// TIA Portal V20 export
FUNCTION_BLOCK "PR_IRVisionCheckSeq_Soft2.0 1_workflow_93eeda"   // FB47, LAD
{ S7_Optimized_Access := 'TRUE' }
// stored: MemoryReserve 100, SetENOAutomatically false
   VAR_INPUT
      iAutoRunning : Bool;
      iFaultReset : Bool;
      iIRMesaureProbeDown : Bool;
      iIRMesaureProbeUp : Bool;
      iIndexCylHome : Bool;
      iIndexProbeOut : Bool;
      iInspectionOver : Bool;
      iManualEntryConfirm : Bool;
      iMesauringOver : Bool;
      iProbeCylHome : Bool;
      iRFIDReadError : Bool;
      iRFIDReadOver : Bool;
      iReject : Bool;
      iReset_fault : Bool;
      iRetry : Bool;
      iRetryCount : Int;
      iSstMode : Bool;
      iSstPB : Bool;
      iStartFrmFibroseq : Bool;
   END_VAR
   VAR_OUTPUT
      qCameraLight : Bool;
      qError : Array[0..9] of Bool;
      qIRProbeDown : Bool;
      qIRProbeUp : Bool;
      qIRVisionCheckOver : Bool;
      qIndexProbeIn : Bool;
      qIndexProbeOut : Bool;
      qMessage : Array[0..9] of Bool;
   END_VAR
   VAR
      c20_ChkRecoveryStatus_T1 : Bool;
      c20_ChkRecoveryStatus_T2 : Bool;
      c20_ChkRecoveryStatus_T3 : Bool;
      c20_ChkRecoveryStatus_T4 : Bool;
      c22_WtRFIDReadOver_T1 : Bool;
      c22_WtRFIDReadOver_T2 : Bool;
      c23_ChkRetryCountOver_T1 : Bool;
      c23_ChkRetryCountOver_T2 : Bool;
      c24_WtOperatorDecisionRead_T1 : Bool;
      c24_WtOperatorDecisionRead_T2 : Bool;
      c25_ChkPartWorkable_T1 : Bool;
      c25_ChkPartWorkable_T2 : Bool;
      c91_WtRFIDWriteOver_T1 : Bool;
      c91_WtRFIDWriteOver_T2 : Bool;
      c92_ChkWriteRetryCountOver_T1 : Bool;
      c92_ChkWriteRetryCountOver_T2 : Bool;
      c93_WtOperatorDecisionWrite_T1 : Bool;
      c93_WtOperatorDecisionWrite_T2 : Bool;
      StateNo : Int;
      s100_WtStartLow : Bool;
      s100_WtStartLow_T1 : Bool;
      s10_WtStartFrmFibroSeq : Bool;
      s10_WtStartFrmFibroSeq_T1 : Bool;
      s1_WtResetRel : Bool;
      s1_WtResetRel_T1 : Bool;
      s20_ChkRecoveryStatus : Bool;
      s20_ChkRecoveryStatus_T1 : Bool;
      s20_ChkRecoveryStatus_T2 : Bool;
      s20_ChkRecoveryStatus_T3 : Bool;
      s20_ChkRecoveryStatus_T4 : Bool;
      s21_WtProbeIndexCylHome : Bool;
      s21_WtProbeIndexCylHome_T1 : Bool;
      s22_WtRFIDReadOver : Bool;
      s22_WtRFIDReadOver_T1 : Bool;
      s22_WtRFIDReadOver_T2 : Bool;
      s23_ChkRetryCountOver : Bool;
      s23_ChkRetryCountOver_T1 : Bool;
      s23_ChkRetryCountOver_T2 : Bool;
      s24_WtOperatorDecisionRead : Bool;
      s24_WtOperatorDecisionRead_T1 : Bool;
      s24_WtOperatorDecisionRead_T2 : Bool;
      s25_ChkPartWorkable : Bool;
      s25_ChkPartWorkable_T1 : Bool;
      s25_ChkPartWorkable_T2 : Bool;
      s30_WtOperatorAck : Bool;
      s30_WtOperatorAck_T1 : Bool;
      s50_WtIRMeasureProbeAtTest : Bool;
      s50_WtIRMeasureProbeAtTest_T1 : Bool;
      s60_WtMeasurementOver : Bool;
      s60_WtMeasurementOver_T1 : Bool;
      s70_WtIRMeasureProbeUp : Bool;
      s70_WtIRMeasureProbeUp_T1 : Bool;
      s80_WtIndexingProbeOut : Bool;
      s80_WtIndexingProbeOut_T1 : Bool;
      s90_WtVisionInspectionOver : Bool;
      s90_WtVisionInspectionOver_T1 : Bool;
      s91_WtRFIDWriteOver : Bool;
      s91_WtRFIDWriteOver_T1 : Bool;
      s91_WtRFIDWriteOver_T2 : Bool;
      s92_ChkWriteRetryCountOver : Bool;
      s92_ChkWriteRetryCountOver_T1 : Bool;
      s92_ChkWriteRetryCountOver_T2 : Bool;
      s93_WtOperatorDecisionWrite : Bool;
      s93_WtOperatorDecisionWrite_T1 : Bool;
      s93_WtOperatorDecisionWrite_T2 : Bool;
      s94_WtAllSystemAtHome : Bool;
      s94_WtAllSystemAtHome_T1 : Bool;
      sAbnormalStatus : Bool;
      sIRInProgress : Bool;
      sPartWorkable : Bool;
      sRFReadRetryCount : Int;
      sRFWriteError : Bool;
      sRFWriteOver : Bool;
      sRFWriteRetryCount : Int;
      sSst : Bool;
      sSstPulse : Bool;
      sSstRise : Bool;
      sStWtResetRel : Bool;
      sStWtResetRel_T1 : Bool;
      sTimeouTime : TON_TIME;
      sVisionInProgress : Bool;
   END_VAR
   VAR_TEMP
      tOne : Bool;
   END_VAR
   VAR_TEMP   // added for the SCL form of the ladder/FBD networks
      _w1 : Bool;
   END_VAR
BEGIN

REGION Network 1
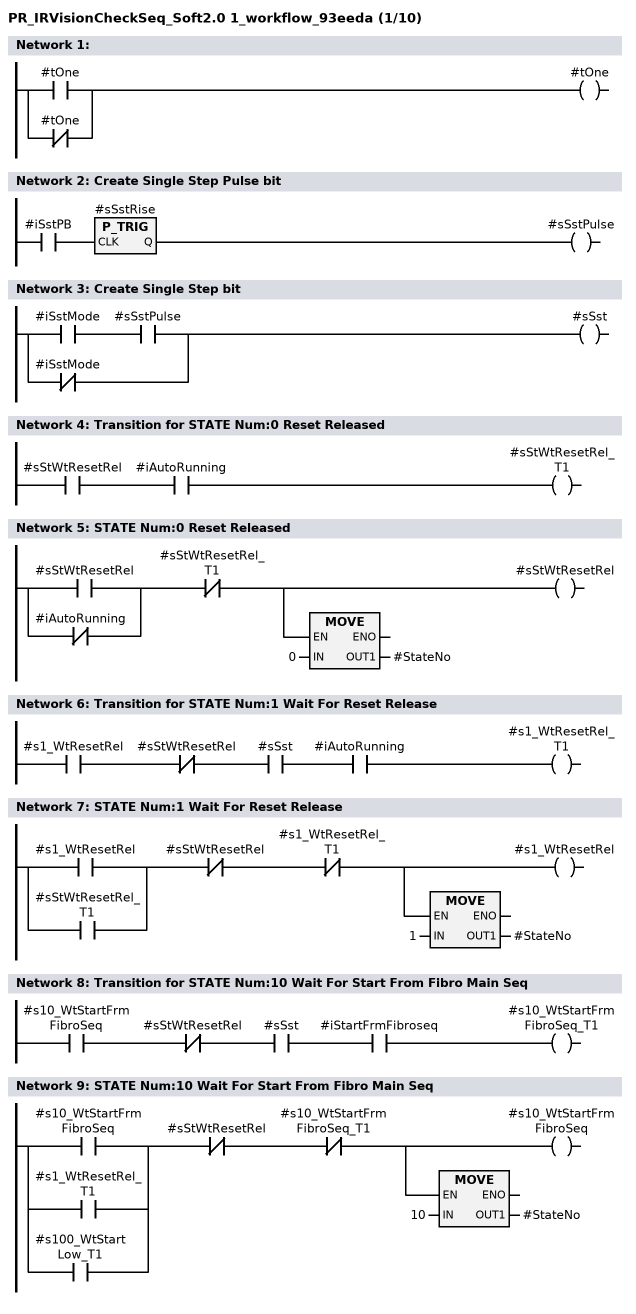
   RUNG wire#powerrail
      Contact( #tOne )
      wire#w1
      Coil( #tOne )
   END_RUNG
   RUNG wire#powerrail
      I_Contact( #tOne )
   END_RUNG wire#w1
   // the same network as SCL:
   #tOne := #tOne OR NOT #tOne;
END_REGION

REGION Network 2: Create Single Step Pulse bit
   RUNG wire#powerrail
      Contact( #iSstPB )
      P_Trig( #sSstRise )
      Coil( #sSstPulse )
   END_RUNG
   // the same network as SCL:
   #_w1 := #iSstPB AND NOT #sSstRise;   // rising edge
   #sSstRise := #iSstPB;
   #sSstPulse := #_w1;
END_REGION

REGION Network 3: Create Single Step bit
   RUNG wire#powerrail
      Contact( #iSstMode )
      Contact( #sSstPulse )
      wire#w1
      Coil( #sSst )
   END_RUNG
   RUNG wire#powerrail
      I_Contact( #iSstMode )
   END_RUNG wire#w1
   // the same network as SCL:
   #sSst := (#iSstMode AND #sSstPulse) OR NOT #iSstMode;
END_REGION

REGION Network 4: Transition for STATE Num:0 Reset Released
   RUNG wire#powerrail
      Contact( #sStWtResetRel )
      Contact( #iAutoRunning )
      Coil( #sStWtResetRel_T1 )
   END_RUNG
   // the same network as SCL:
   #sStWtResetRel_T1 := #sStWtResetRel AND #iAutoRunning;
END_REGION

REGION Network 5: STATE Num:0 Reset Released
   RUNG wire#powerrail
      Contact( #sStWtResetRel )
      wire#w1
      I_Contact( #sStWtResetRel_T1 )
      wire#w2
      Coil( #sStWtResetRel )
   END_RUNG
   RUNG wire#powerrail
      I_Contact( #iAutoRunning )
   END_RUNG wire#w1
   RUNG wire#w2
      { S7_GenerateENO := "TRUE" } Move(in := 0, out1 => #StateNo)
   END_RUNG
   // the same network as SCL:
   #sStWtResetRel := (#sStWtResetRel OR NOT #iAutoRunning) AND NOT #sStWtResetRel_T1;
   IF #sStWtResetRel THEN #StateNo := 0; END_IF;
END_REGION

REGION Network 6: Transition for STATE Num:1 Wait For Reset Release
   RUNG wire#powerrail
      Contact( #s1_WtResetRel )
      I_Contact( #sStWtResetRel )
      Contact( #sSst )
      Contact( #iAutoRunning )
      Coil( #s1_WtResetRel_T1 )
   END_RUNG
   // the same network as SCL:
   #s1_WtResetRel_T1 := #s1_WtResetRel AND NOT #sStWtResetRel AND #sSst AND #iAutoRunning;
END_REGION

REGION Network 7: STATE Num:1 Wait For Reset Release
   RUNG wire#powerrail
      Contact( #s1_WtResetRel )
      wire#w1
      I_Contact( #sStWtResetRel )
      I_Contact( #s1_WtResetRel_T1 )
      wire#w2
      Coil( #s1_WtResetRel )
   END_RUNG
   RUNG wire#powerrail
      Contact( #sStWtResetRel_T1 )
   END_RUNG wire#w1
   RUNG wire#w2
      { S7_GenerateENO := "TRUE" } Move(in := 1, out1 => #StateNo)
   END_RUNG
   // the same network as SCL:
   #s1_WtResetRel := (#s1_WtResetRel OR #sStWtResetRel_T1) AND NOT #sStWtResetRel AND NOT #s1_WtResetRel_T1;
   IF #s1_WtResetRel THEN #StateNo := 1; END_IF;
END_REGION

REGION Network 8: Transition for STATE Num:10 Wait For Start From Fibro Main Seq
   RUNG wire#powerrail
      Contact( #s10_WtStartFrmFibroSeq )
      I_Contact( #sStWtResetRel )
      Contact( #sSst )
      Contact( #iStartFrmFibroseq )
      Coil( #s10_WtStartFrmFibroSeq_T1 )
   END_RUNG
   // the same network as SCL:
   #s10_WtStartFrmFibroSeq_T1 := #s10_WtStartFrmFibroSeq AND NOT #sStWtResetRel AND #sSst AND #iStartFrmFibroseq;
END_REGION

REGION Network 9: STATE Num:10 Wait For Start From Fibro Main Seq
   RUNG wire#powerrail
      Contact( #s10_WtStartFrmFibroSeq )
      wire#w1
      I_Contact( #sStWtResetRel )
      I_Contact( #s10_WtStartFrmFibroSeq_T1 )
      wire#w2
      Coil( #s10_WtStartFrmFibroSeq )
   END_RUNG
   RUNG wire#powerrail
      Contact( #s1_WtResetRel_T1 )
   END_RUNG wire#w1
   RUNG wire#powerrail
      Contact( #s100_WtStartLow_T1 )
   END_RUNG wire#w1
   RUNG wire#w2
      { S7_GenerateENO := "TRUE" } Move(in := 10, out1 => #StateNo)
   END_RUNG
   // the same network as SCL:
   #s10_WtStartFrmFibroSeq := (#s10_WtStartFrmFibroSeq OR #s1_WtResetRel_T1 OR #s100_WtStartLow_T1) AND NOT #sStWtResetRel AND NOT #s10_WtStartFrmFibroSeq_T1;
   IF #s10_WtStartFrmFibroSeq THEN #StateNo := 10; END_IF;
END_REGION

REGION Network 10: Actions for STATE Num:10 Wait For Start From Fibro Main Seq
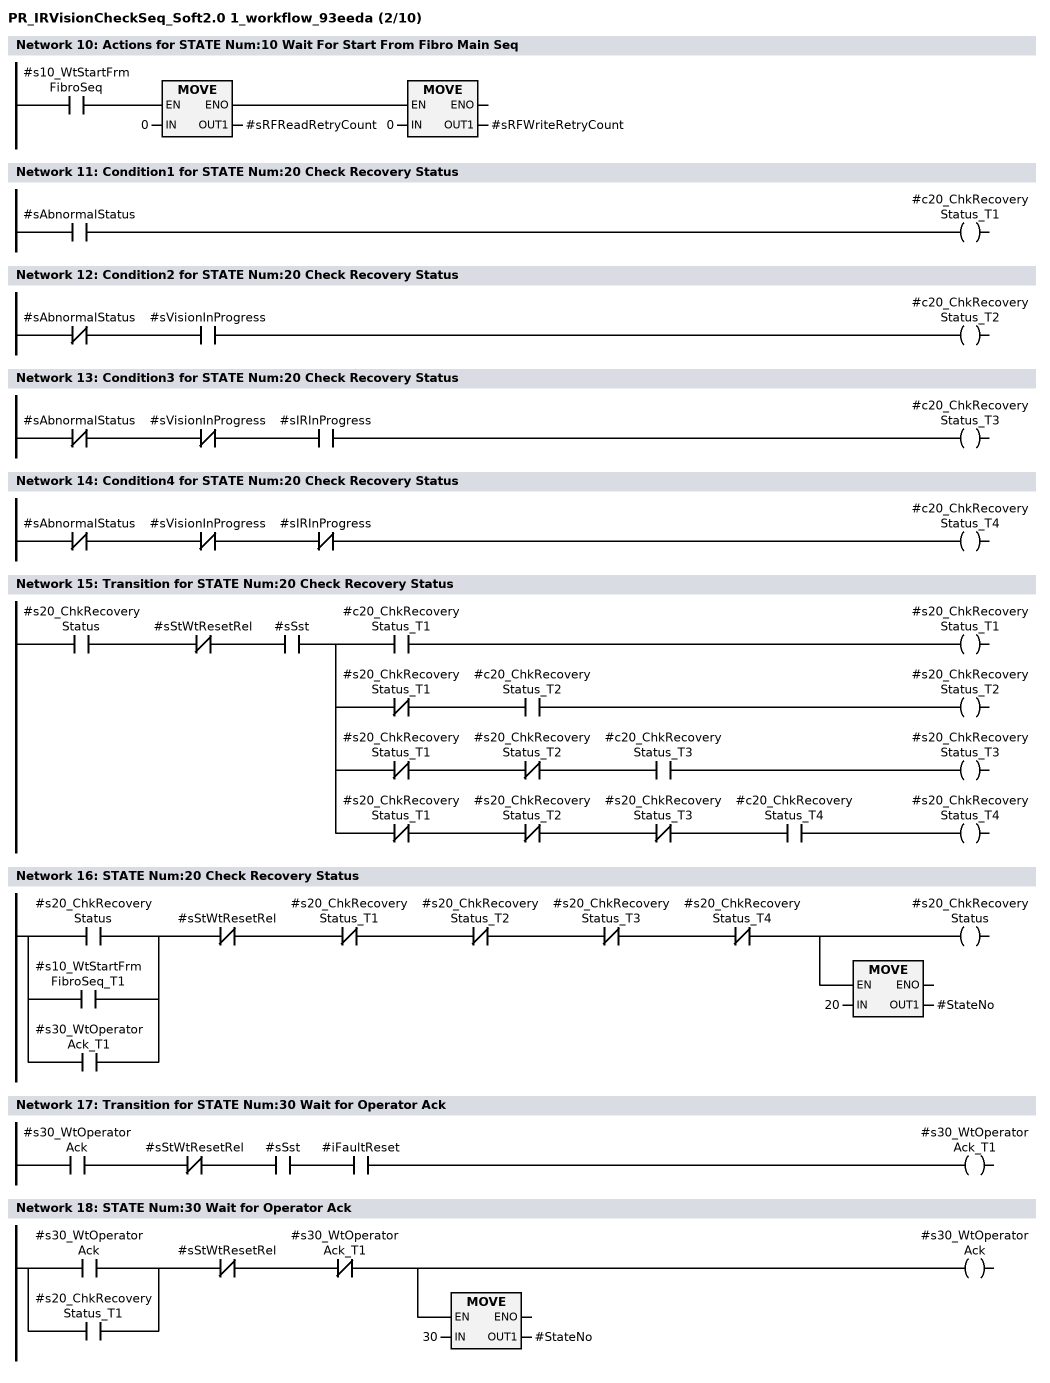
   RUNG wire#powerrail
      Contact( #s10_WtStartFrmFibroSeq )
      Move(in := 0, out1 => #sRFReadRetryCount)
      Move(in := 0, out1 => #sRFWriteRetryCount)
   END_RUNG
   // the same network as SCL:
   IF #s10_WtStartFrmFibroSeq THEN
       #sRFReadRetryCount := 0;
       #sRFWriteRetryCount := 0;
   END_IF;
END_REGION

REGION Network 11: Condition1 for STATE Num:20 Check Recovery Status
   RUNG wire#powerrail
      Contact( #sAbnormalStatus )
      Coil( #c20_ChkRecoveryStatus_T1 )
   END_RUNG
   // the same network as SCL:
   #c20_ChkRecoveryStatus_T1 := #sAbnormalStatus;
END_REGION

REGION Network 12: Condition2 for STATE Num:20 Check Recovery Status
   RUNG wire#powerrail
      I_Contact( #sAbnormalStatus )
      Contact( #sVisionInProgress )
      Coil( #c20_ChkRecoveryStatus_T2 )
   END_RUNG
   // the same network as SCL:
   #c20_ChkRecoveryStatus_T2 := NOT #sAbnormalStatus AND #sVisionInProgress;
END_REGION

REGION Network 13: Condition3 for STATE Num:20 Check Recovery Status
   RUNG wire#powerrail
      I_Contact( #sAbnormalStatus )
      I_Contact( #sVisionInProgress )
      Contact( #sIRInProgress )
      Coil( #c20_ChkRecoveryStatus_T3 )
   END_RUNG
   // the same network as SCL:
   #c20_ChkRecoveryStatus_T3 := NOT #sAbnormalStatus AND NOT #sVisionInProgress AND #sIRInProgress;
END_REGION

REGION Network 14: Condition4 for STATE Num:20 Check Recovery Status
   RUNG wire#powerrail
      I_Contact( #sAbnormalStatus )
      I_Contact( #sVisionInProgress )
      I_Contact( #sIRInProgress )
      Coil( #c20_ChkRecoveryStatus_T4 )
   END_RUNG
   // the same network as SCL:
   #c20_ChkRecoveryStatus_T4 := NOT #sAbnormalStatus AND NOT #sVisionInProgress AND NOT #sIRInProgress;
END_REGION

REGION Network 15: Transition for STATE Num:20 Check Recovery Status
   RUNG wire#powerrail
      Contact( #s20_ChkRecoveryStatus )
      I_Contact( #sStWtResetRel )
      Contact( #sSst )
      wire#w1
      Contact( #c20_ChkRecoveryStatus_T1 )
      Coil( #s20_ChkRecoveryStatus_T1 )
   END_RUNG
   RUNG wire#w1
      I_Contact( #s20_ChkRecoveryStatus_T1 )
      Contact( #c20_ChkRecoveryStatus_T2 )
      Coil( #s20_ChkRecoveryStatus_T2 )
   END_RUNG
   RUNG wire#w1
      I_Contact( #s20_ChkRecoveryStatus_T1 )
      I_Contact( #s20_ChkRecoveryStatus_T2 )
      Contact( #c20_ChkRecoveryStatus_T3 )
      Coil( #s20_ChkRecoveryStatus_T3 )
   END_RUNG
   RUNG wire#w1
      I_Contact( #s20_ChkRecoveryStatus_T1 )
      I_Contact( #s20_ChkRecoveryStatus_T2 )
      I_Contact( #s20_ChkRecoveryStatus_T3 )
      Contact( #c20_ChkRecoveryStatus_T4 )
      Coil( #s20_ChkRecoveryStatus_T4 )
   END_RUNG
   // the same network as SCL:
   #_w1 := #s20_ChkRecoveryStatus AND NOT #sStWtResetRel AND #sSst;
   #s20_ChkRecoveryStatus_T1 := #_w1 AND #c20_ChkRecoveryStatus_T1;
   #s20_ChkRecoveryStatus_T2 := #_w1 AND NOT #s20_ChkRecoveryStatus_T1 AND #c20_ChkRecoveryStatus_T2;
   #s20_ChkRecoveryStatus_T3 := #_w1 AND NOT #s20_ChkRecoveryStatus_T1 AND NOT #s20_ChkRecoveryStatus_T2 AND #c20_ChkRecoveryStatus_T3;
   #s20_ChkRecoveryStatus_T4 := #_w1 AND NOT #s20_ChkRecoveryStatus_T1 AND NOT #s20_ChkRecoveryStatus_T2 AND NOT #s20_ChkRecoveryStatus_T3 AND #c20_ChkRecoveryStatus_T4;
END_REGION

REGION Network 16: STATE Num:20 Check Recovery Status
   RUNG wire#powerrail
      Contact( #s20_ChkRecoveryStatus )
      wire#w1
      I_Contact( #sStWtResetRel )
      I_Contact( #s20_ChkRecoveryStatus_T1 )
      I_Contact( #s20_ChkRecoveryStatus_T2 )
      I_Contact( #s20_ChkRecoveryStatus_T3 )
      I_Contact( #s20_ChkRecoveryStatus_T4 )
      wire#w2
      Coil( #s20_ChkRecoveryStatus )
   END_RUNG
   RUNG wire#powerrail
      Contact( #s10_WtStartFrmFibroSeq_T1 )
   END_RUNG wire#w1
   RUNG wire#powerrail
      Contact( #s30_WtOperatorAck_T1 )
   END_RUNG wire#w1
   RUNG wire#w2
      { S7_GenerateENO := "TRUE" } Move(in := 20, out1 => #StateNo)
   END_RUNG
   // the same network as SCL:
   #s20_ChkRecoveryStatus := (#s20_ChkRecoveryStatus OR #s10_WtStartFrmFibroSeq_T1 OR #s30_WtOperatorAck_T1) AND NOT #sStWtResetRel AND NOT #s20_ChkRecoveryStatus_T1 AND NOT #s20_ChkRecoveryStatus_T2 AND NOT #s20_ChkRecoveryStatus_T3 AND NOT #s20_ChkRecoveryStatus_T4;
   IF #s20_ChkRecoveryStatus THEN #StateNo := 20; END_IF;
END_REGION

REGION Network 17: Transition for STATE Num:30 Wait for Operator Ack
   RUNG wire#powerrail
      Contact( #s30_WtOperatorAck )
      I_Contact( #sStWtResetRel )
      Contact( #sSst )
      Contact( #iFaultReset )
      Coil( #s30_WtOperatorAck_T1 )
   END_RUNG
   // the same network as SCL:
   #s30_WtOperatorAck_T1 := #s30_WtOperatorAck AND NOT #sStWtResetRel AND #sSst AND #iFaultReset;
END_REGION

REGION Network 18: STATE Num:30 Wait for Operator Ack
   RUNG wire#powerrail
      Contact( #s30_WtOperatorAck )
      wire#w1
      I_Contact( #sStWtResetRel )
      I_Contact( #s30_WtOperatorAck_T1 )
      wire#w2
      Coil( #s30_WtOperatorAck )
   END_RUNG
   RUNG wire#powerrail
      Contact( #s20_ChkRecoveryStatus_T1 )
   END_RUNG wire#w1
   RUNG wire#w2
      { S7_GenerateENO := "TRUE" } Move(in := 30, out1 => #StateNo)
   END_RUNG
   // the same network as SCL:
   #s30_WtOperatorAck := (#s30_WtOperatorAck OR #s20_ChkRecoveryStatus_T1) AND NOT #sStWtResetRel AND NOT #s30_WtOperatorAck_T1;
   IF #s30_WtOperatorAck THEN #StateNo := 30; END_IF;
END_REGION

REGION Network 19: Actions for STATE Num:30 Wait for Operator Ack
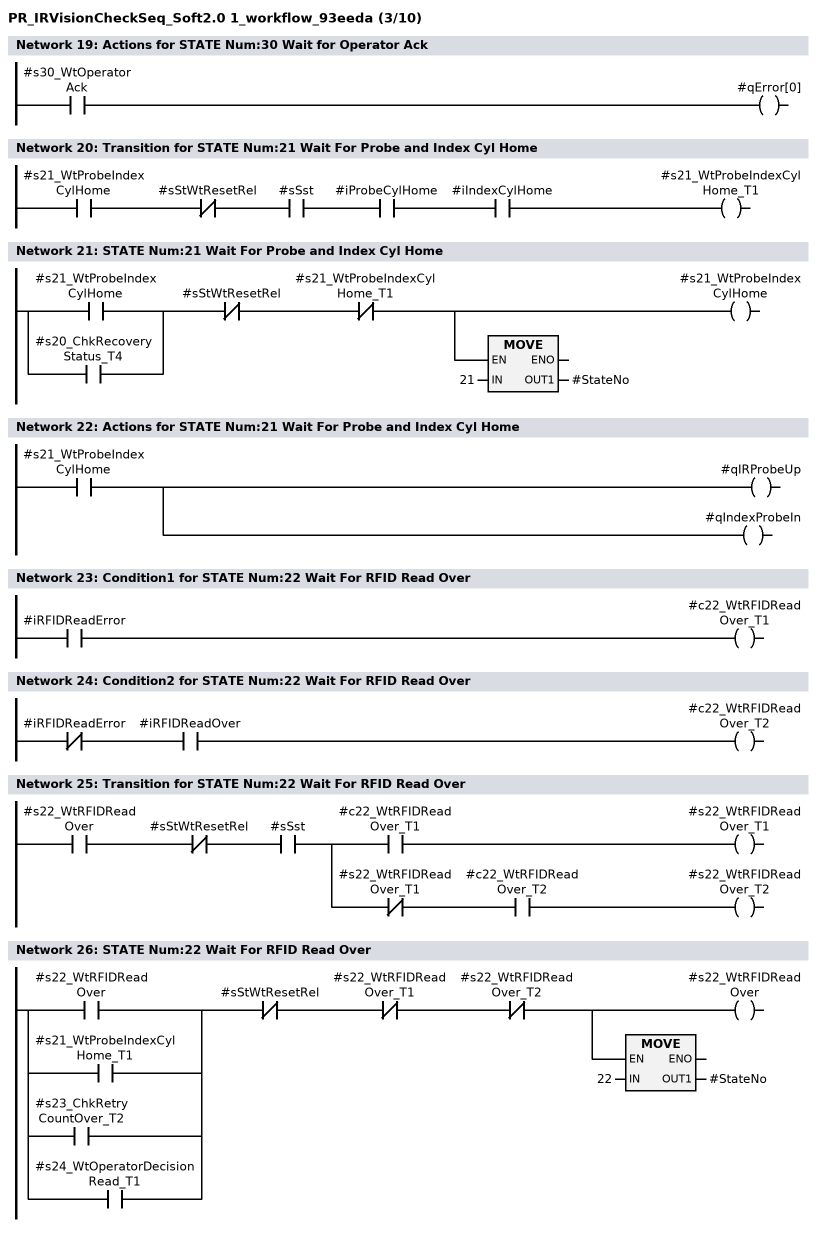
   RUNG wire#powerrail
      Contact( #s30_WtOperatorAck )
      Coil( #qError[0] )
   END_RUNG
   // the same network as SCL:
   #qError[0] := #s30_WtOperatorAck;
END_REGION

REGION Network 20: Transition for STATE Num:21 Wait For Probe and Index Cyl Home
   RUNG wire#powerrail
      Contact( #s21_WtProbeIndexCylHome )
      I_Contact( #sStWtResetRel )
      Contact( #sSst )
      Contact( #iProbeCylHome )
      Contact( #iIndexCylHome )
      Coil( #s21_WtProbeIndexCylHome_T1 )
   END_RUNG
   // the same network as SCL:
   #s21_WtProbeIndexCylHome_T1 := #s21_WtProbeIndexCylHome AND NOT #sStWtResetRel AND #sSst AND #iProbeCylHome AND #iIndexCylHome;
END_REGION

REGION Network 21: STATE Num:21 Wait For Probe and Index Cyl Home
   RUNG wire#powerrail
      Contact( #s21_WtProbeIndexCylHome )
      wire#w1
      I_Contact( #sStWtResetRel )
      I_Contact( #s21_WtProbeIndexCylHome_T1 )
      wire#w2
      Coil( #s21_WtProbeIndexCylHome )
   END_RUNG
   RUNG wire#powerrail
      Contact( #s20_ChkRecoveryStatus_T4 )
   END_RUNG wire#w1
   RUNG wire#w2
      { S7_GenerateENO := "TRUE" } Move(in := 21, out1 => #StateNo)
   END_RUNG
   // the same network as SCL:
   #s21_WtProbeIndexCylHome := (#s21_WtProbeIndexCylHome OR #s20_ChkRecoveryStatus_T4) AND NOT #sStWtResetRel AND NOT #s21_WtProbeIndexCylHome_T1;
   IF #s21_WtProbeIndexCylHome THEN #StateNo := 21; END_IF;
END_REGION

REGION Network 22: Actions for STATE Num:21 Wait For Probe and Index Cyl Home
   RUNG wire#powerrail
      Contact( #s21_WtProbeIndexCylHome )
      wire#w1
      Coil( #qIRProbeUp )
   END_RUNG
   RUNG wire#w1
      Coil( #qIndexProbeIn )
   END_RUNG
   // the same network as SCL:
   #qIRProbeUp := #s21_WtProbeIndexCylHome;
   #qIndexProbeIn := #s21_WtProbeIndexCylHome;
END_REGION

REGION Network 23: Condition1 for STATE Num:22 Wait For RFID Read Over
   RUNG wire#powerrail
      Contact( #iRFIDReadError )
      Coil( #c22_WtRFIDReadOver_T1 )
   END_RUNG
   // the same network as SCL:
   #c22_WtRFIDReadOver_T1 := #iRFIDReadError;
END_REGION

REGION Network 24: Condition2 for STATE Num:22 Wait For RFID Read Over
   RUNG wire#powerrail
      I_Contact( #iRFIDReadError )
      Contact( #iRFIDReadOver )
      Coil( #c22_WtRFIDReadOver_T2 )
   END_RUNG
   // the same network as SCL:
   #c22_WtRFIDReadOver_T2 := NOT #iRFIDReadError AND #iRFIDReadOver;
END_REGION

REGION Network 25: Transition for STATE Num:22 Wait For RFID Read Over
   RUNG wire#powerrail
      Contact( #s22_WtRFIDReadOver )
      I_Contact( #sStWtResetRel )
      Contact( #sSst )
      wire#w1
      Contact( #c22_WtRFIDReadOver_T1 )
      Coil( #s22_WtRFIDReadOver_T1 )
   END_RUNG
   RUNG wire#w1
      I_Contact( #s22_WtRFIDReadOver_T1 )
      Contact( #c22_WtRFIDReadOver_T2 )
      Coil( #s22_WtRFIDReadOver_T2 )
   END_RUNG
   // the same network as SCL:
   #_w1 := #s22_WtRFIDReadOver AND NOT #sStWtResetRel AND #sSst;
   #s22_WtRFIDReadOver_T1 := #_w1 AND #c22_WtRFIDReadOver_T1;
   #s22_WtRFIDReadOver_T2 := #_w1 AND NOT #s22_WtRFIDReadOver_T1 AND #c22_WtRFIDReadOver_T2;
END_REGION

REGION Network 26: STATE Num:22 Wait For RFID Read Over
   RUNG wire#powerrail
      Contact( #s22_WtRFIDReadOver )
      wire#w1
      I_Contact( #sStWtResetRel )
      I_Contact( #s22_WtRFIDReadOver_T1 )
      I_Contact( #s22_WtRFIDReadOver_T2 )
      wire#w2
      Coil( #s22_WtRFIDReadOver )
   END_RUNG
   RUNG wire#powerrail
      Contact( #s21_WtProbeIndexCylHome_T1 )
   END_RUNG wire#w1
   RUNG wire#powerrail
      Contact( #s23_ChkRetryCountOver_T2 )
   END_RUNG wire#w1
   RUNG wire#powerrail
      Contact( #s24_WtOperatorDecisionRead_T1 )
   END_RUNG wire#w1
   RUNG wire#w2
      { S7_GenerateENO := "TRUE" } Move(in := 22, out1 => #StateNo)
   END_RUNG
   // the same network as SCL:
   #s22_WtRFIDReadOver := (#s22_WtRFIDReadOver OR #s21_WtProbeIndexCylHome_T1 OR #s23_ChkRetryCountOver_T2 OR #s24_WtOperatorDecisionRead_T1) AND NOT #sStWtResetRel AND NOT #s22_WtRFIDReadOver_T1 AND NOT #s22_WtRFIDReadOver_T2;
   IF #s22_WtRFIDReadOver THEN #StateNo := 22; END_IF;
END_REGION

REGION Network 27: Transition Actions T1 for STATE Num:22 Wait For RFID Read Over
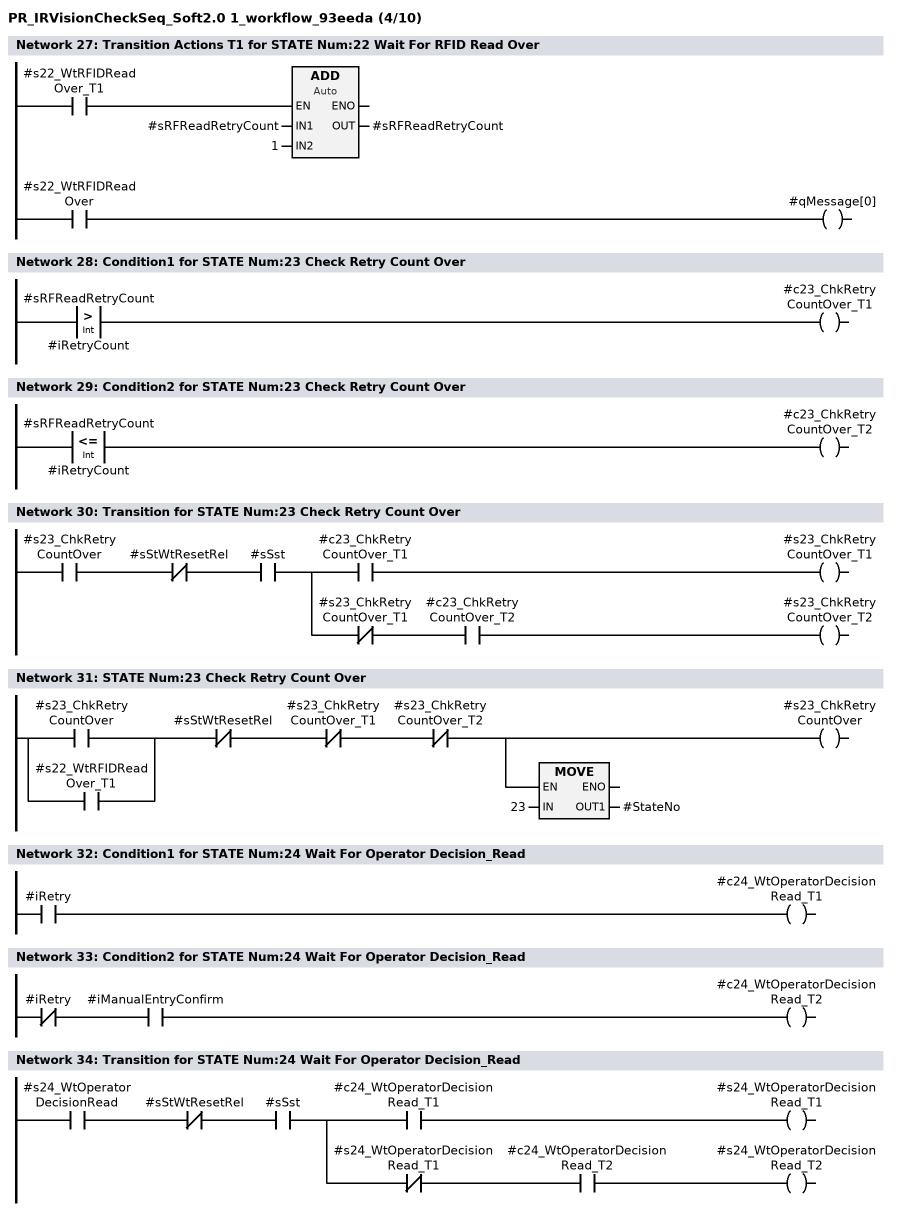
   RUNG wire#powerrail
      Contact( #s22_WtRFIDReadOver_T1 )
      Add(in1 := #sRFReadRetryCount, in2 := 1, out => #sRFReadRetryCount)
   END_RUNG
   RUNG wire#powerrail
      Contact( #s22_WtRFIDReadOver )
      Coil( #qMessage[0] )
   END_RUNG
   // the same network as SCL:
   IF #s22_WtRFIDReadOver_T1 THEN #sRFReadRetryCount := #sRFReadRetryCount + 1; END_IF;
   #qMessage[0] := #s22_WtRFIDReadOver;
END_REGION

REGION Network 28: Condition1 for STATE Num:23 Check Retry Count Over
   RUNG wire#powerrail
      { S7_Templates := "SrcType := Int" } GT_Contact(in1 := #sRFReadRetryCount, in2 := #iRetryCount)
      Coil( #c23_ChkRetryCountOver_T1 )
   END_RUNG
   // the same network as SCL:
   #c23_ChkRetryCountOver_T1 := #sRFReadRetryCount > #iRetryCount;
END_REGION

REGION Network 29: Condition2 for STATE Num:23 Check Retry Count Over
   RUNG wire#powerrail
      { S7_Templates := "SrcType := Int" } LE_Contact(in1 := #sRFReadRetryCount, in2 := #iRetryCount)
      Coil( #c23_ChkRetryCountOver_T2 )
   END_RUNG
   // the same network as SCL:
   #c23_ChkRetryCountOver_T2 := #sRFReadRetryCount <= #iRetryCount;
END_REGION

REGION Network 30: Transition for STATE Num:23 Check Retry Count Over
   RUNG wire#powerrail
      Contact( #s23_ChkRetryCountOver )
      I_Contact( #sStWtResetRel )
      Contact( #sSst )
      wire#w1
      Contact( #c23_ChkRetryCountOver_T1 )
      Coil( #s23_ChkRetryCountOver_T1 )
   END_RUNG
   RUNG wire#w1
      I_Contact( #s23_ChkRetryCountOver_T1 )
      Contact( #c23_ChkRetryCountOver_T2 )
      Coil( #s23_ChkRetryCountOver_T2 )
   END_RUNG
   // the same network as SCL:
   #_w1 := #s23_ChkRetryCountOver AND NOT #sStWtResetRel AND #sSst;
   #s23_ChkRetryCountOver_T1 := #_w1 AND #c23_ChkRetryCountOver_T1;
   #s23_ChkRetryCountOver_T2 := #_w1 AND NOT #s23_ChkRetryCountOver_T1 AND #c23_ChkRetryCountOver_T2;
END_REGION

REGION Network 31: STATE Num:23 Check Retry Count Over
   RUNG wire#powerrail
      Contact( #s23_ChkRetryCountOver )
      wire#w1
      I_Contact( #sStWtResetRel )
      I_Contact( #s23_ChkRetryCountOver_T1 )
      I_Contact( #s23_ChkRetryCountOver_T2 )
      wire#w2
      Coil( #s23_ChkRetryCountOver )
   END_RUNG
   RUNG wire#powerrail
      Contact( #s22_WtRFIDReadOver_T1 )
   END_RUNG wire#w1
   RUNG wire#w2
      { S7_GenerateENO := "TRUE" } Move(in := 23, out1 => #StateNo)
   END_RUNG
   // the same network as SCL:
   #s23_ChkRetryCountOver := (#s23_ChkRetryCountOver OR #s22_WtRFIDReadOver_T1) AND NOT #sStWtResetRel AND NOT #s23_ChkRetryCountOver_T1 AND NOT #s23_ChkRetryCountOver_T2;
   IF #s23_ChkRetryCountOver THEN #StateNo := 23; END_IF;
END_REGION

REGION Network 32: Condition1 for STATE Num:24 Wait For Operator Decision_Read
   RUNG wire#powerrail
      Contact( #iRetry )
      Coil( #c24_WtOperatorDecisionRead_T1 )
   END_RUNG
   // the same network as SCL:
   #c24_WtOperatorDecisionRead_T1 := #iRetry;
END_REGION

REGION Network 33: Condition2 for STATE Num:24 Wait For Operator Decision_Read
   RUNG wire#powerrail
      I_Contact( #iRetry )
      Contact( #iManualEntryConfirm )
      Coil( #c24_WtOperatorDecisionRead_T2 )
   END_RUNG
   // the same network as SCL:
   #c24_WtOperatorDecisionRead_T2 := NOT #iRetry AND #iManualEntryConfirm;
END_REGION

REGION Network 34: Transition for STATE Num:24 Wait For Operator Decision_Read
   RUNG wire#powerrail
      Contact( #s24_WtOperatorDecisionRead )
      I_Contact( #sStWtResetRel )
      Contact( #sSst )
      wire#w1
      Contact( #c24_WtOperatorDecisionRead_T1 )
      Coil( #s24_WtOperatorDecisionRead_T1 )
   END_RUNG
   RUNG wire#w1
      I_Contact( #s24_WtOperatorDecisionRead_T1 )
      Contact( #c24_WtOperatorDecisionRead_T2 )
      Coil( #s24_WtOperatorDecisionRead_T2 )
   END_RUNG
   // the same network as SCL:
   #_w1 := #s24_WtOperatorDecisionRead AND NOT #sStWtResetRel AND #sSst;
   #s24_WtOperatorDecisionRead_T1 := #_w1 AND #c24_WtOperatorDecisionRead_T1;
   #s24_WtOperatorDecisionRead_T2 := #_w1 AND NOT #s24_WtOperatorDecisionRead_T1 AND #c24_WtOperatorDecisionRead_T2;
END_REGION

REGION Network 35: STATE Num:24 Wait For Operator Decision_Read
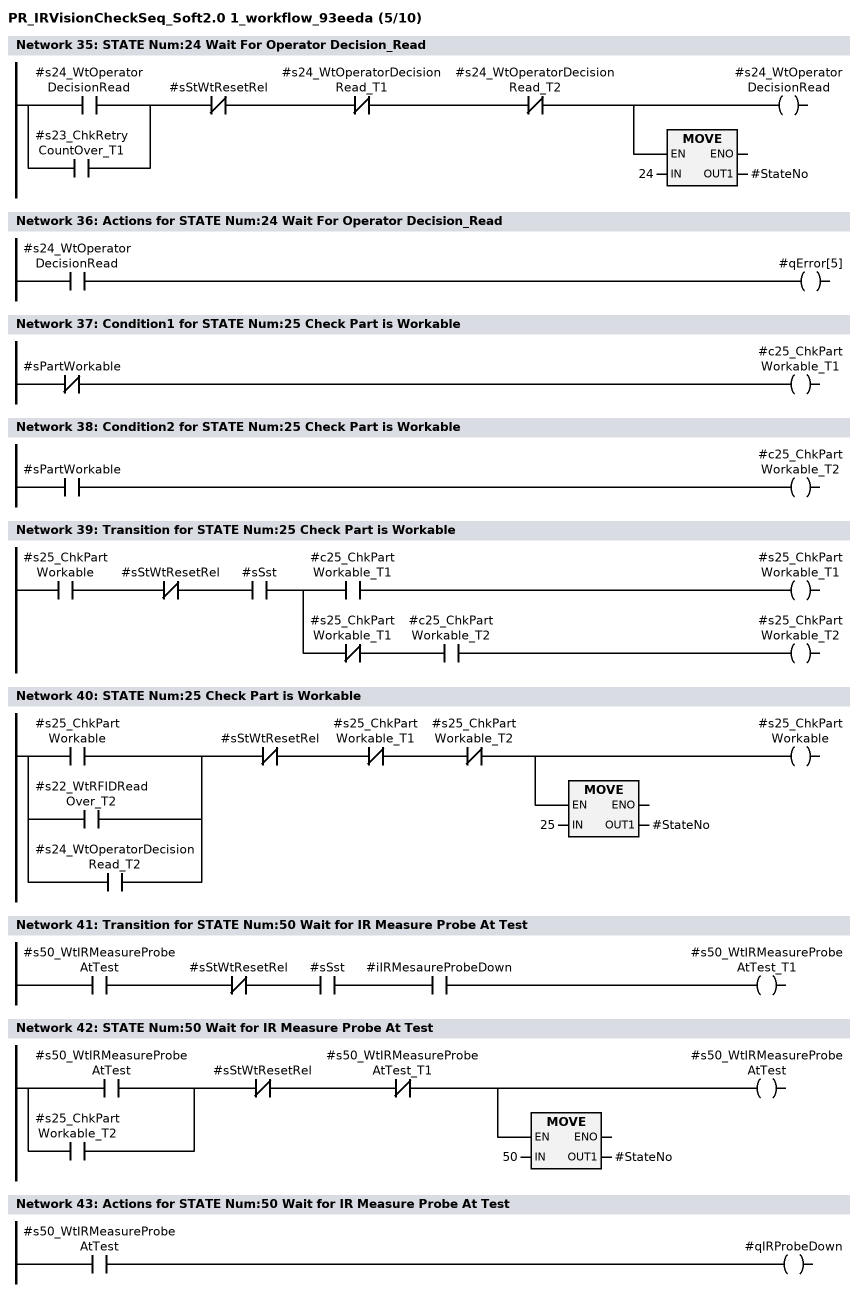
   RUNG wire#powerrail
      Contact( #s24_WtOperatorDecisionRead )
      wire#w1
      I_Contact( #sStWtResetRel )
      I_Contact( #s24_WtOperatorDecisionRead_T1 )
      I_Contact( #s24_WtOperatorDecisionRead_T2 )
      wire#w2
      Coil( #s24_WtOperatorDecisionRead )
   END_RUNG
   RUNG wire#powerrail
      Contact( #s23_ChkRetryCountOver_T1 )
   END_RUNG wire#w1
   RUNG wire#w2
      { S7_GenerateENO := "TRUE" } Move(in := 24, out1 => #StateNo)
   END_RUNG
   // the same network as SCL:
   #s24_WtOperatorDecisionRead := (#s24_WtOperatorDecisionRead OR #s23_ChkRetryCountOver_T1) AND NOT #sStWtResetRel AND NOT #s24_WtOperatorDecisionRead_T1 AND NOT #s24_WtOperatorDecisionRead_T2;
   IF #s24_WtOperatorDecisionRead THEN #StateNo := 24; END_IF;
END_REGION

REGION Network 36: Actions for STATE Num:24 Wait For Operator Decision_Read
   RUNG wire#powerrail
      Contact( #s24_WtOperatorDecisionRead )
      Coil( #qError[5] )
   END_RUNG
   // the same network as SCL:
   #qError[5] := #s24_WtOperatorDecisionRead;
END_REGION

REGION Network 37: Condition1 for STATE Num:25 Check Part is Workable
   RUNG wire#powerrail
      I_Contact( #sPartWorkable )
      Coil( #c25_ChkPartWorkable_T1 )
   END_RUNG
   // the same network as SCL:
   #c25_ChkPartWorkable_T1 := NOT #sPartWorkable;
END_REGION

REGION Network 38: Condition2 for STATE Num:25 Check Part is Workable
   RUNG wire#powerrail
      Contact( #sPartWorkable )
      Coil( #c25_ChkPartWorkable_T2 )
   END_RUNG
   // the same network as SCL:
   #c25_ChkPartWorkable_T2 := #sPartWorkable;
END_REGION

REGION Network 39: Transition for STATE Num:25 Check Part is Workable
   RUNG wire#powerrail
      Contact( #s25_ChkPartWorkable )
      I_Contact( #sStWtResetRel )
      Contact( #sSst )
      wire#w1
      Contact( #c25_ChkPartWorkable_T1 )
      Coil( #s25_ChkPartWorkable_T1 )
   END_RUNG
   RUNG wire#w1
      I_Contact( #s25_ChkPartWorkable_T1 )
      Contact( #c25_ChkPartWorkable_T2 )
      Coil( #s25_ChkPartWorkable_T2 )
   END_RUNG
   // the same network as SCL:
   #_w1 := #s25_ChkPartWorkable AND NOT #sStWtResetRel AND #sSst;
   #s25_ChkPartWorkable_T1 := #_w1 AND #c25_ChkPartWorkable_T1;
   #s25_ChkPartWorkable_T2 := #_w1 AND NOT #s25_ChkPartWorkable_T1 AND #c25_ChkPartWorkable_T2;
END_REGION

REGION Network 40: STATE Num:25 Check Part is Workable
   RUNG wire#powerrail
      Contact( #s25_ChkPartWorkable )
      wire#w1
      I_Contact( #sStWtResetRel )
      I_Contact( #s25_ChkPartWorkable_T1 )
      I_Contact( #s25_ChkPartWorkable_T2 )
      wire#w2
      Coil( #s25_ChkPartWorkable )
   END_RUNG
   RUNG wire#powerrail
      Contact( #s22_WtRFIDReadOver_T2 )
   END_RUNG wire#w1
   RUNG wire#powerrail
      Contact( #s24_WtOperatorDecisionRead_T2 )
   END_RUNG wire#w1
   RUNG wire#w2
      { S7_GenerateENO := "TRUE" } Move(in := 25, out1 => #StateNo)
   END_RUNG
   // the same network as SCL:
   #s25_ChkPartWorkable := (#s25_ChkPartWorkable OR #s22_WtRFIDReadOver_T2 OR #s24_WtOperatorDecisionRead_T2) AND NOT #sStWtResetRel AND NOT #s25_ChkPartWorkable_T1 AND NOT #s25_ChkPartWorkable_T2;
   IF #s25_ChkPartWorkable THEN #StateNo := 25; END_IF;
END_REGION

REGION Network 41: Transition for STATE Num:50 Wait for IR Measure Probe At Test
   RUNG wire#powerrail
      Contact( #s50_WtIRMeasureProbeAtTest )
      I_Contact( #sStWtResetRel )
      Contact( #sSst )
      Contact( #iIRMesaureProbeDown )
      Coil( #s50_WtIRMeasureProbeAtTest_T1 )
   END_RUNG
   // the same network as SCL:
   #s50_WtIRMeasureProbeAtTest_T1 := #s50_WtIRMeasureProbeAtTest AND NOT #sStWtResetRel AND #sSst AND #iIRMesaureProbeDown;
END_REGION

REGION Network 42: STATE Num:50 Wait for IR Measure Probe At Test
   RUNG wire#powerrail
      Contact( #s50_WtIRMeasureProbeAtTest )
      wire#w1
      I_Contact( #sStWtResetRel )
      I_Contact( #s50_WtIRMeasureProbeAtTest_T1 )
      wire#w2
      Coil( #s50_WtIRMeasureProbeAtTest )
   END_RUNG
   RUNG wire#powerrail
      Contact( #s25_ChkPartWorkable_T2 )
   END_RUNG wire#w1
   RUNG wire#w2
      { S7_GenerateENO := "TRUE" } Move(in := 50, out1 => #StateNo)
   END_RUNG
   // the same network as SCL:
   #s50_WtIRMeasureProbeAtTest := (#s50_WtIRMeasureProbeAtTest OR #s25_ChkPartWorkable_T2) AND NOT #sStWtResetRel AND NOT #s50_WtIRMeasureProbeAtTest_T1;
   IF #s50_WtIRMeasureProbeAtTest THEN #StateNo := 50; END_IF;
END_REGION

REGION Network 43: Actions for STATE Num:50 Wait for IR Measure Probe At Test
   RUNG wire#powerrail
      Contact( #s50_WtIRMeasureProbeAtTest )
      Coil( #qIRProbeDown )
   END_RUNG
   // the same network as SCL:
   #qIRProbeDown := #s50_WtIRMeasureProbeAtTest;
END_REGION

REGION Network 44: Transition for STATE Num:60 Wait For Measurement Over
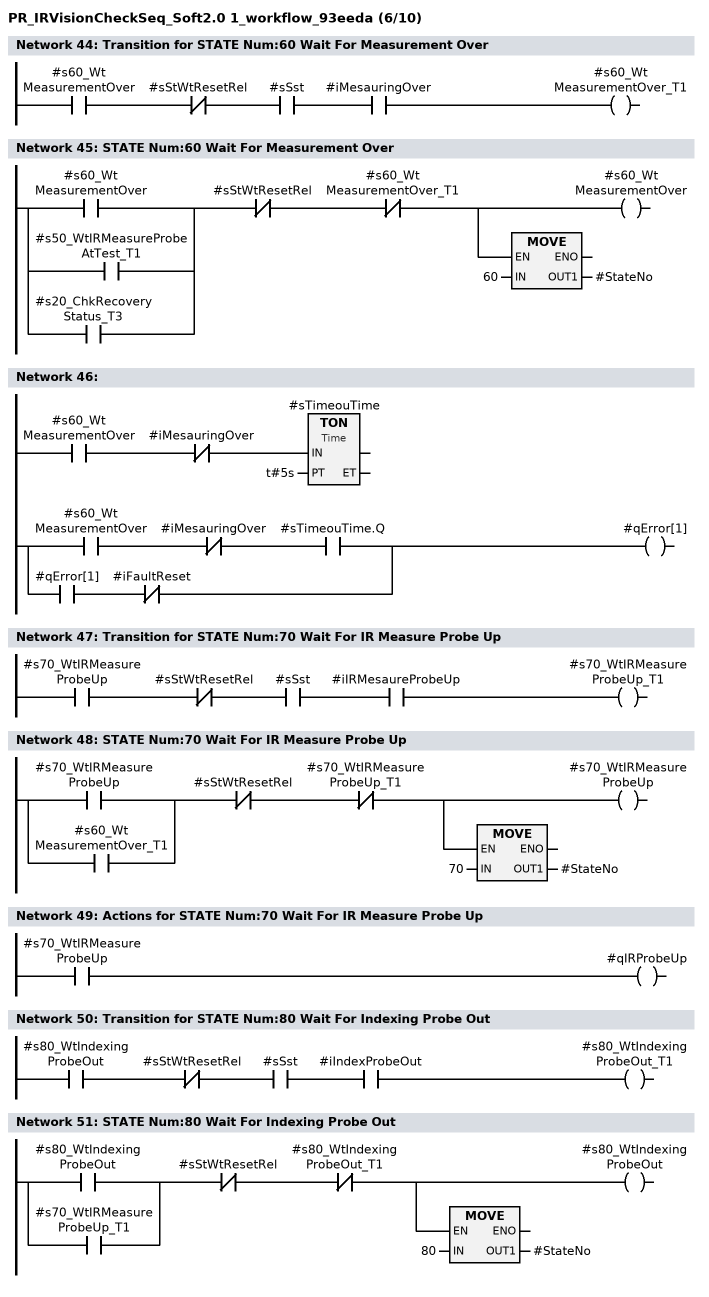
   RUNG wire#powerrail
      Contact( #s60_WtMeasurementOver )
      I_Contact( #sStWtResetRel )
      Contact( #sSst )
      Contact( #iMesauringOver )
      Coil( #s60_WtMeasurementOver_T1 )
   END_RUNG
   // the same network as SCL:
   #s60_WtMeasurementOver_T1 := #s60_WtMeasurementOver AND NOT #sStWtResetRel AND #sSst AND #iMesauringOver;
END_REGION

REGION Network 45: STATE Num:60 Wait For Measurement Over
   RUNG wire#powerrail
      Contact( #s60_WtMeasurementOver )
      wire#w1
      I_Contact( #sStWtResetRel )
      I_Contact( #s60_WtMeasurementOver_T1 )
      wire#w2
      Coil( #s60_WtMeasurementOver )
   END_RUNG
   RUNG wire#powerrail
      Contact( #s50_WtIRMeasureProbeAtTest_T1 )
   END_RUNG wire#w1
   RUNG wire#powerrail
      Contact( #s20_ChkRecoveryStatus_T3 )
   END_RUNG wire#w1
   RUNG wire#w2
      { S7_GenerateENO := "TRUE" } Move(in := 60, out1 => #StateNo)
   END_RUNG
   // the same network as SCL:
   #s60_WtMeasurementOver := (#s60_WtMeasurementOver OR #s50_WtIRMeasureProbeAtTest_T1 OR #s20_ChkRecoveryStatus_T3) AND NOT #sStWtResetRel AND NOT #s60_WtMeasurementOver_T1;
   IF #s60_WtMeasurementOver THEN #StateNo := 60; END_IF;
END_REGION

REGION Network 46
   RUNG wire#powerrail
      Contact( #s60_WtMeasurementOver )
      I_Contact( #iMesauringOver )
      { S7_Templates := "time_type := Time" } #sTimeouTime.TON(pt := t#5s, et =>)
   END_RUNG
   RUNG wire#powerrail
      Contact( #s60_WtMeasurementOver )
      I_Contact( #iMesauringOver )
      Contact( #sTimeouTime.Q )
      wire#w1
      Coil( #qError[1] )
   END_RUNG
   RUNG wire#powerrail
      Contact( #qError[1] )
      I_Contact( #iFaultReset )
   END_RUNG wire#w1
   // the same network as SCL:
   #sTimeouTime(IN := #s60_WtMeasurementOver AND NOT #iMesauringOver, PT := t#5s);   // TON
   #qError[1] := (#s60_WtMeasurementOver AND NOT #iMesauringOver AND #sTimeouTime.Q) OR (#qError[1] AND NOT #iFaultReset);
END_REGION

REGION Network 47: Transition for STATE Num:70 Wait For IR Measure Probe Up
   RUNG wire#powerrail
      Contact( #s70_WtIRMeasureProbeUp )
      I_Contact( #sStWtResetRel )
      Contact( #sSst )
      Contact( #iIRMesaureProbeUp )
      Coil( #s70_WtIRMeasureProbeUp_T1 )
   END_RUNG
   // the same network as SCL:
   #s70_WtIRMeasureProbeUp_T1 := #s70_WtIRMeasureProbeUp AND NOT #sStWtResetRel AND #sSst AND #iIRMesaureProbeUp;
END_REGION

REGION Network 48: STATE Num:70 Wait For IR Measure Probe Up
   RUNG wire#powerrail
      Contact( #s70_WtIRMeasureProbeUp )
      wire#w1
      I_Contact( #sStWtResetRel )
      I_Contact( #s70_WtIRMeasureProbeUp_T1 )
      wire#w2
      Coil( #s70_WtIRMeasureProbeUp )
   END_RUNG
   RUNG wire#powerrail
      Contact( #s60_WtMeasurementOver_T1 )
   END_RUNG wire#w1
   RUNG wire#w2
      { S7_GenerateENO := "TRUE" } Move(in := 70, out1 => #StateNo)
   END_RUNG
   // the same network as SCL:
   #s70_WtIRMeasureProbeUp := (#s70_WtIRMeasureProbeUp OR #s60_WtMeasurementOver_T1) AND NOT #sStWtResetRel AND NOT #s70_WtIRMeasureProbeUp_T1;
   IF #s70_WtIRMeasureProbeUp THEN #StateNo := 70; END_IF;
END_REGION

REGION Network 49: Actions for STATE Num:70 Wait For IR Measure Probe Up
   RUNG wire#powerrail
      Contact( #s70_WtIRMeasureProbeUp )
      Coil( #qIRProbeUp )
   END_RUNG
   // the same network as SCL:
   #qIRProbeUp := #s70_WtIRMeasureProbeUp;
END_REGION

REGION Network 50: Transition for STATE Num:80 Wait For Indexing Probe Out
   RUNG wire#powerrail
      Contact( #s80_WtIndexingProbeOut )
      I_Contact( #sStWtResetRel )
      Contact( #sSst )
      Contact( #iIndexProbeOut )
      Coil( #s80_WtIndexingProbeOut_T1 )
   END_RUNG
   // the same network as SCL:
   #s80_WtIndexingProbeOut_T1 := #s80_WtIndexingProbeOut AND NOT #sStWtResetRel AND #sSst AND #iIndexProbeOut;
END_REGION

REGION Network 51: STATE Num:80 Wait For Indexing Probe Out
   RUNG wire#powerrail
      Contact( #s80_WtIndexingProbeOut )
      wire#w1
      I_Contact( #sStWtResetRel )
      I_Contact( #s80_WtIndexingProbeOut_T1 )
      wire#w2
      Coil( #s80_WtIndexingProbeOut )
   END_RUNG
   RUNG wire#powerrail
      Contact( #s70_WtIRMeasureProbeUp_T1 )
   END_RUNG wire#w1
   RUNG wire#w2
      { S7_GenerateENO := "TRUE" } Move(in := 80, out1 => #StateNo)
   END_RUNG
   // the same network as SCL:
   #s80_WtIndexingProbeOut := (#s80_WtIndexingProbeOut OR #s70_WtIRMeasureProbeUp_T1) AND NOT #sStWtResetRel AND NOT #s80_WtIndexingProbeOut_T1;
   IF #s80_WtIndexingProbeOut THEN #StateNo := 80; END_IF;
END_REGION

REGION Network 52: Actions for STATE Num:80 Wait For Indexing Probe Out
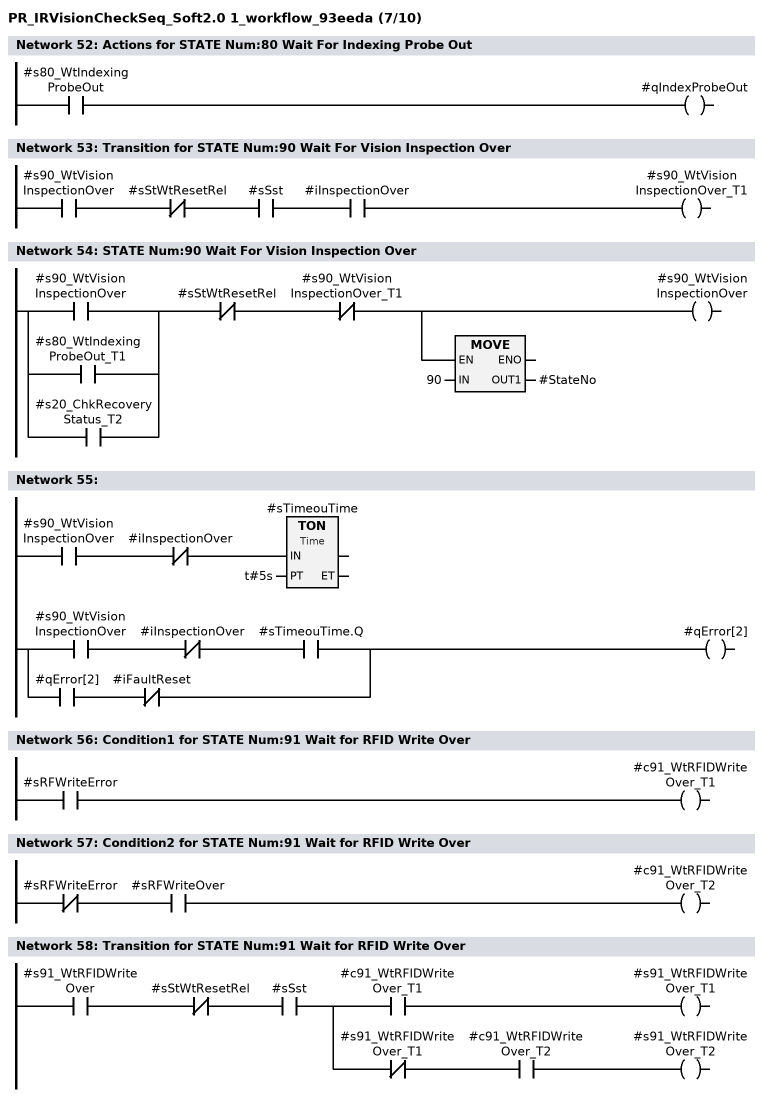
   RUNG wire#powerrail
      Contact( #s80_WtIndexingProbeOut )
      Coil( #qIndexProbeOut )
   END_RUNG
   // the same network as SCL:
   #qIndexProbeOut := #s80_WtIndexingProbeOut;
END_REGION

REGION Network 53: Transition for STATE Num:90 Wait For Vision Inspection Over
   RUNG wire#powerrail
      Contact( #s90_WtVisionInspectionOver )
      I_Contact( #sStWtResetRel )
      Contact( #sSst )
      Contact( #iInspectionOver )
      Coil( #s90_WtVisionInspectionOver_T1 )
   END_RUNG
   // the same network as SCL:
   #s90_WtVisionInspectionOver_T1 := #s90_WtVisionInspectionOver AND NOT #sStWtResetRel AND #sSst AND #iInspectionOver;
END_REGION

REGION Network 54: STATE Num:90 Wait For Vision Inspection Over
   RUNG wire#powerrail
      Contact( #s90_WtVisionInspectionOver )
      wire#w1
      I_Contact( #sStWtResetRel )
      I_Contact( #s90_WtVisionInspectionOver_T1 )
      wire#w2
      Coil( #s90_WtVisionInspectionOver )
   END_RUNG
   RUNG wire#powerrail
      Contact( #s80_WtIndexingProbeOut_T1 )
   END_RUNG wire#w1
   RUNG wire#powerrail
      Contact( #s20_ChkRecoveryStatus_T2 )
   END_RUNG wire#w1
   RUNG wire#w2
      { S7_GenerateENO := "TRUE" } Move(in := 90, out1 => #StateNo)
   END_RUNG
   // the same network as SCL:
   #s90_WtVisionInspectionOver := (#s90_WtVisionInspectionOver OR #s80_WtIndexingProbeOut_T1 OR #s20_ChkRecoveryStatus_T2) AND NOT #sStWtResetRel AND NOT #s90_WtVisionInspectionOver_T1;
   IF #s90_WtVisionInspectionOver THEN #StateNo := 90; END_IF;
END_REGION

REGION Network 55
   RUNG wire#powerrail
      Contact( #s90_WtVisionInspectionOver )
      I_Contact( #iInspectionOver )
      { S7_Templates := "time_type := Time" } #sTimeouTime.TON(pt := t#5s, et =>)
   END_RUNG
   RUNG wire#powerrail
      Contact( #s90_WtVisionInspectionOver )
      I_Contact( #iInspectionOver )
      Contact( #sTimeouTime.Q )
      wire#w1
      Coil( #qError[2] )
   END_RUNG
   RUNG wire#powerrail
      Contact( #qError[2] )
      I_Contact( #iFaultReset )
   END_RUNG wire#w1
   // the same network as SCL:
   #sTimeouTime(IN := #s90_WtVisionInspectionOver AND NOT #iInspectionOver, PT := t#5s);   // TON
   #qError[2] := (#s90_WtVisionInspectionOver AND NOT #iInspectionOver AND #sTimeouTime.Q) OR (#qError[2] AND NOT #iFaultReset);
END_REGION

REGION Network 56: Condition1 for STATE Num:91 Wait for RFID Write Over
   RUNG wire#powerrail
      Contact( #sRFWriteError )
      Coil( #c91_WtRFIDWriteOver_T1 )
   END_RUNG
   // the same network as SCL:
   #c91_WtRFIDWriteOver_T1 := #sRFWriteError;
END_REGION

REGION Network 57: Condition2 for STATE Num:91 Wait for RFID Write Over
   RUNG wire#powerrail
      I_Contact( #sRFWriteError )
      Contact( #sRFWriteOver )
      Coil( #c91_WtRFIDWriteOver_T2 )
   END_RUNG
   // the same network as SCL:
   #c91_WtRFIDWriteOver_T2 := NOT #sRFWriteError AND #sRFWriteOver;
END_REGION

REGION Network 58: Transition for STATE Num:91 Wait for RFID Write Over
   RUNG wire#powerrail
      Contact( #s91_WtRFIDWriteOver )
      I_Contact( #sStWtResetRel )
      Contact( #sSst )
      wire#w1
      Contact( #c91_WtRFIDWriteOver_T1 )
      Coil( #s91_WtRFIDWriteOver_T1 )
   END_RUNG
   RUNG wire#w1
      I_Contact( #s91_WtRFIDWriteOver_T1 )
      Contact( #c91_WtRFIDWriteOver_T2 )
      Coil( #s91_WtRFIDWriteOver_T2 )
   END_RUNG
   // the same network as SCL:
   #_w1 := #s91_WtRFIDWriteOver AND NOT #sStWtResetRel AND #sSst;
   #s91_WtRFIDWriteOver_T1 := #_w1 AND #c91_WtRFIDWriteOver_T1;
   #s91_WtRFIDWriteOver_T2 := #_w1 AND NOT #s91_WtRFIDWriteOver_T1 AND #c91_WtRFIDWriteOver_T2;
END_REGION

REGION Network 59: STATE Num:91 Wait for RFID Write Over
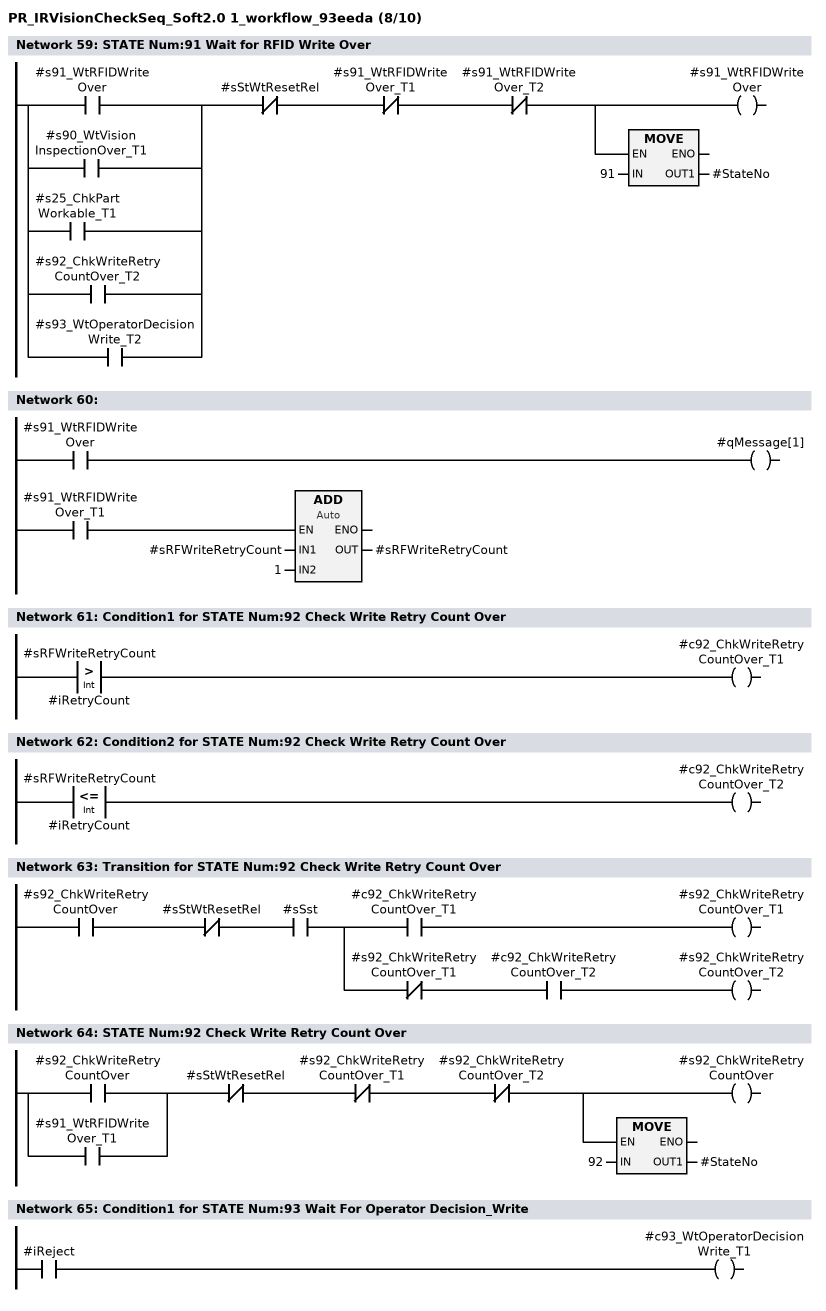
   RUNG wire#powerrail
      Contact( #s91_WtRFIDWriteOver )
      wire#w1
      I_Contact( #sStWtResetRel )
      I_Contact( #s91_WtRFIDWriteOver_T1 )
      I_Contact( #s91_WtRFIDWriteOver_T2 )
      wire#w2
      Coil( #s91_WtRFIDWriteOver )
   END_RUNG
   RUNG wire#powerrail
      Contact( #s90_WtVisionInspectionOver_T1 )
   END_RUNG wire#w1
   RUNG wire#powerrail
      Contact( #s25_ChkPartWorkable_T1 )
   END_RUNG wire#w1
   RUNG wire#powerrail
      Contact( #s92_ChkWriteRetryCountOver_T2 )
   END_RUNG wire#w1
   RUNG wire#powerrail
      Contact( #s93_WtOperatorDecisionWrite_T2 )
   END_RUNG wire#w1
   RUNG wire#w2
      { S7_GenerateENO := "TRUE" } Move(in := 91, out1 => #StateNo)
   END_RUNG
   // the same network as SCL:
   #s91_WtRFIDWriteOver := (#s91_WtRFIDWriteOver OR #s90_WtVisionInspectionOver_T1 OR #s25_ChkPartWorkable_T1 OR #s92_ChkWriteRetryCountOver_T2 OR #s93_WtOperatorDecisionWrite_T2) AND NOT #sStWtResetRel AND NOT #s91_WtRFIDWriteOver_T1 AND NOT #s91_WtRFIDWriteOver_T2;
   IF #s91_WtRFIDWriteOver THEN #StateNo := 91; END_IF;
END_REGION

REGION Network 60
   RUNG wire#powerrail
      Contact( #s91_WtRFIDWriteOver )
      Coil( #qMessage[1] )
   END_RUNG
   RUNG wire#powerrail
      Contact( #s91_WtRFIDWriteOver_T1 )
      Add(in1 := #sRFWriteRetryCount, in2 := 1, out => #sRFWriteRetryCount)
   END_RUNG
   // the same network as SCL:
   #qMessage[1] := #s91_WtRFIDWriteOver;
   IF #s91_WtRFIDWriteOver_T1 THEN #sRFWriteRetryCount := #sRFWriteRetryCount + 1; END_IF;
END_REGION

REGION Network 61: Condition1 for STATE Num:92 Check Write Retry Count Over
   RUNG wire#powerrail
      { S7_Templates := "SrcType := Int" } GT_Contact(in1 := #sRFWriteRetryCount, in2 := #iRetryCount)
      Coil( #c92_ChkWriteRetryCountOver_T1 )
   END_RUNG
   // the same network as SCL:
   #c92_ChkWriteRetryCountOver_T1 := #sRFWriteRetryCount > #iRetryCount;
END_REGION

REGION Network 62: Condition2 for STATE Num:92 Check Write Retry Count Over
   RUNG wire#powerrail
      { S7_Templates := "SrcType := Int" } LE_Contact(in1 := #sRFWriteRetryCount, in2 := #iRetryCount)
      Coil( #c92_ChkWriteRetryCountOver_T2 )
   END_RUNG
   // the same network as SCL:
   #c92_ChkWriteRetryCountOver_T2 := #sRFWriteRetryCount <= #iRetryCount;
END_REGION

REGION Network 63: Transition for STATE Num:92 Check Write Retry Count Over
   RUNG wire#powerrail
      Contact( #s92_ChkWriteRetryCountOver )
      I_Contact( #sStWtResetRel )
      Contact( #sSst )
      wire#w1
      Contact( #c92_ChkWriteRetryCountOver_T1 )
      Coil( #s92_ChkWriteRetryCountOver_T1 )
   END_RUNG
   RUNG wire#w1
      I_Contact( #s92_ChkWriteRetryCountOver_T1 )
      Contact( #c92_ChkWriteRetryCountOver_T2 )
      Coil( #s92_ChkWriteRetryCountOver_T2 )
   END_RUNG
   // the same network as SCL:
   #_w1 := #s92_ChkWriteRetryCountOver AND NOT #sStWtResetRel AND #sSst;
   #s92_ChkWriteRetryCountOver_T1 := #_w1 AND #c92_ChkWriteRetryCountOver_T1;
   #s92_ChkWriteRetryCountOver_T2 := #_w1 AND NOT #s92_ChkWriteRetryCountOver_T1 AND #c92_ChkWriteRetryCountOver_T2;
END_REGION

REGION Network 64: STATE Num:92 Check Write Retry Count Over
   RUNG wire#powerrail
      Contact( #s92_ChkWriteRetryCountOver )
      wire#w1
      I_Contact( #sStWtResetRel )
      I_Contact( #s92_ChkWriteRetryCountOver_T1 )
      I_Contact( #s92_ChkWriteRetryCountOver_T2 )
      wire#w2
      Coil( #s92_ChkWriteRetryCountOver )
   END_RUNG
   RUNG wire#powerrail
      Contact( #s91_WtRFIDWriteOver_T1 )
   END_RUNG wire#w1
   RUNG wire#w2
      { S7_GenerateENO := "TRUE" } Move(in := 92, out1 => #StateNo)
   END_RUNG
   // the same network as SCL:
   #s92_ChkWriteRetryCountOver := (#s92_ChkWriteRetryCountOver OR #s91_WtRFIDWriteOver_T1) AND NOT #sStWtResetRel AND NOT #s92_ChkWriteRetryCountOver_T1 AND NOT #s92_ChkWriteRetryCountOver_T2;
   IF #s92_ChkWriteRetryCountOver THEN #StateNo := 92; END_IF;
END_REGION

REGION Network 65: Condition1 for STATE Num:93 Wait For Operator Decision_Write
   RUNG wire#powerrail
      Contact( #iReject )
      Coil( #c93_WtOperatorDecisionWrite_T1 )
   END_RUNG
   // the same network as SCL:
   #c93_WtOperatorDecisionWrite_T1 := #iReject;
END_REGION

REGION Network 66: Condition2 for STATE Num:93 Wait For Operator Decision_Write
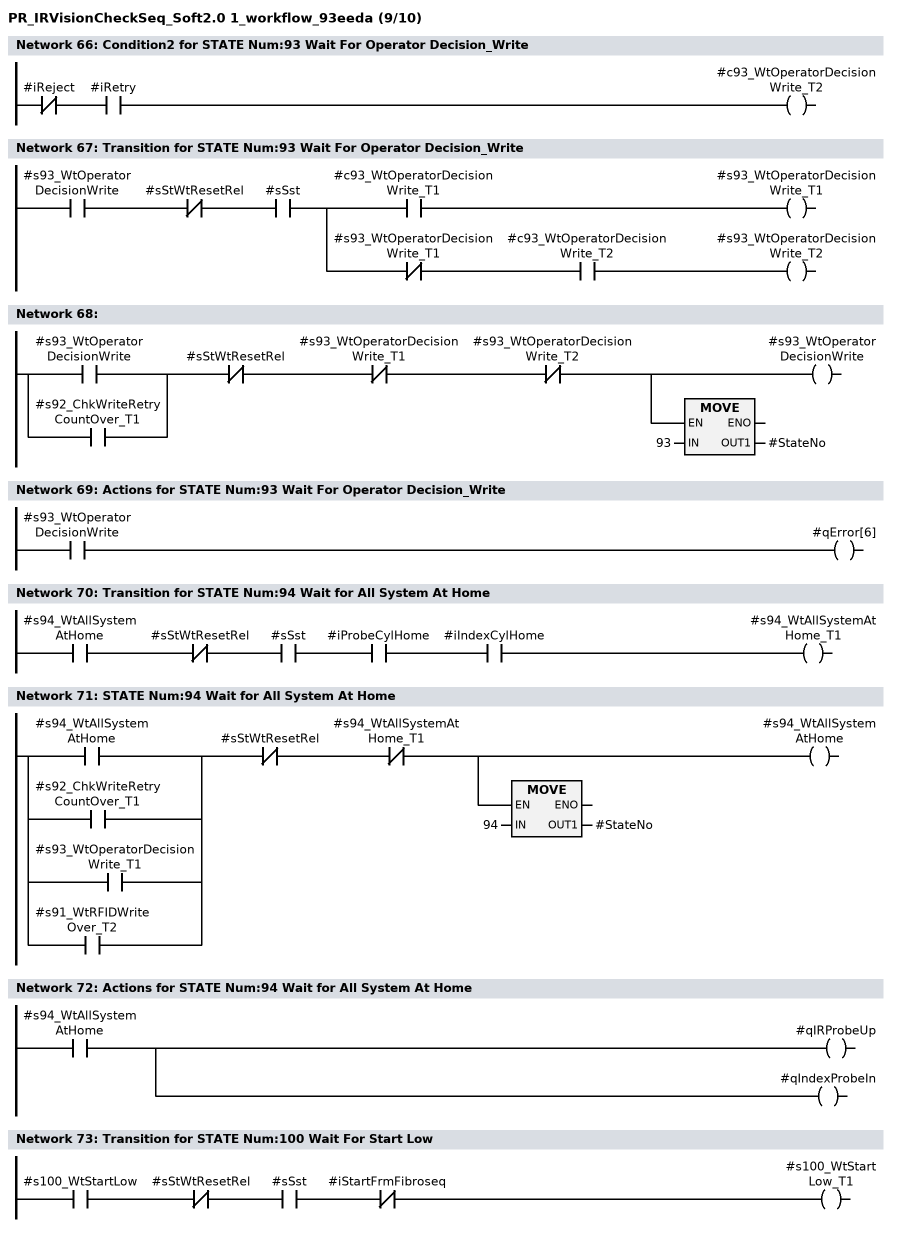
   RUNG wire#powerrail
      I_Contact( #iReject )
      Contact( #iRetry )
      Coil( #c93_WtOperatorDecisionWrite_T2 )
   END_RUNG
   // the same network as SCL:
   #c93_WtOperatorDecisionWrite_T2 := NOT #iReject AND #iRetry;
END_REGION

REGION Network 67: Transition for STATE Num:93 Wait For Operator Decision_Write
   RUNG wire#powerrail
      Contact( #s93_WtOperatorDecisionWrite )
      I_Contact( #sStWtResetRel )
      Contact( #sSst )
      wire#w1
      Contact( #c93_WtOperatorDecisionWrite_T1 )
      Coil( #s93_WtOperatorDecisionWrite_T1 )
   END_RUNG
   RUNG wire#w1
      I_Contact( #s93_WtOperatorDecisionWrite_T1 )
      Contact( #c93_WtOperatorDecisionWrite_T2 )
      Coil( #s93_WtOperatorDecisionWrite_T2 )
   END_RUNG
   // the same network as SCL:
   #_w1 := #s93_WtOperatorDecisionWrite AND NOT #sStWtResetRel AND #sSst;
   #s93_WtOperatorDecisionWrite_T1 := #_w1 AND #c93_WtOperatorDecisionWrite_T1;
   #s93_WtOperatorDecisionWrite_T2 := #_w1 AND NOT #s93_WtOperatorDecisionWrite_T1 AND #c93_WtOperatorDecisionWrite_T2;
END_REGION

REGION Network 68
   RUNG wire#powerrail
      Contact( #s93_WtOperatorDecisionWrite )
      wire#w1
      I_Contact( #sStWtResetRel )
      I_Contact( #s93_WtOperatorDecisionWrite_T1 )
      I_Contact( #s93_WtOperatorDecisionWrite_T2 )
      wire#w2
      Coil( #s93_WtOperatorDecisionWrite )
   END_RUNG
   RUNG wire#powerrail
      Contact( #s92_ChkWriteRetryCountOver_T1 )
   END_RUNG wire#w1
   RUNG wire#w2
      { S7_GenerateENO := "TRUE" } Move(in := 93, out1 => #StateNo)
   END_RUNG
   // the same network as SCL:
   #s93_WtOperatorDecisionWrite := (#s93_WtOperatorDecisionWrite OR #s92_ChkWriteRetryCountOver_T1) AND NOT #sStWtResetRel AND NOT #s93_WtOperatorDecisionWrite_T1 AND NOT #s93_WtOperatorDecisionWrite_T2;
   IF #s93_WtOperatorDecisionWrite THEN #StateNo := 93; END_IF;
END_REGION

REGION Network 69: Actions for STATE Num:93 Wait For Operator Decision_Write
   RUNG wire#powerrail
      Contact( #s93_WtOperatorDecisionWrite )
      Coil( #qError[6] )
   END_RUNG
   // the same network as SCL:
   #qError[6] := #s93_WtOperatorDecisionWrite;
END_REGION

REGION Network 70: Transition for STATE Num:94 Wait for All System At Home
   RUNG wire#powerrail
      Contact( #s94_WtAllSystemAtHome )
      I_Contact( #sStWtResetRel )
      Contact( #sSst )
      Contact( #iProbeCylHome )
      Contact( #iIndexCylHome )
      Coil( #s94_WtAllSystemAtHome_T1 )
   END_RUNG
   // the same network as SCL:
   #s94_WtAllSystemAtHome_T1 := #s94_WtAllSystemAtHome AND NOT #sStWtResetRel AND #sSst AND #iProbeCylHome AND #iIndexCylHome;
END_REGION

REGION Network 71: STATE Num:94 Wait for All System At Home
   RUNG wire#powerrail
      Contact( #s94_WtAllSystemAtHome )
      wire#w1
      I_Contact( #sStWtResetRel )
      I_Contact( #s94_WtAllSystemAtHome_T1 )
      wire#w2
      Coil( #s94_WtAllSystemAtHome )
   END_RUNG
   RUNG wire#powerrail
      Contact( #s92_ChkWriteRetryCountOver_T1 )
   END_RUNG wire#w1
   RUNG wire#powerrail
      Contact( #s93_WtOperatorDecisionWrite_T1 )
   END_RUNG wire#w1
   RUNG wire#powerrail
      Contact( #s91_WtRFIDWriteOver_T2 )
   END_RUNG wire#w1
   RUNG wire#w2
      { S7_GenerateENO := "TRUE" } Move(in := 94, out1 => #StateNo)
   END_RUNG
   // the same network as SCL:
   #s94_WtAllSystemAtHome := (#s94_WtAllSystemAtHome OR #s92_ChkWriteRetryCountOver_T1 OR #s93_WtOperatorDecisionWrite_T1 OR #s91_WtRFIDWriteOver_T2) AND NOT #sStWtResetRel AND NOT #s94_WtAllSystemAtHome_T1;
   IF #s94_WtAllSystemAtHome THEN #StateNo := 94; END_IF;
END_REGION

REGION Network 72: Actions for STATE Num:94 Wait for All System At Home
   RUNG wire#powerrail
      Contact( #s94_WtAllSystemAtHome )
      wire#w1
      Coil( #qIRProbeUp )
   END_RUNG
   RUNG wire#w1
      Coil( #qIndexProbeIn )
   END_RUNG
   // the same network as SCL:
   #qIRProbeUp := #s94_WtAllSystemAtHome;
   #qIndexProbeIn := #s94_WtAllSystemAtHome;
END_REGION

REGION Network 73: Transition for STATE Num:100 Wait For Start Low
   RUNG wire#powerrail
      Contact( #s100_WtStartLow )
      I_Contact( #sStWtResetRel )
      Contact( #sSst )
      I_Contact( #iStartFrmFibroseq )
      Coil( #s100_WtStartLow_T1 )
   END_RUNG
   // the same network as SCL:
   #s100_WtStartLow_T1 := #s100_WtStartLow AND NOT #sStWtResetRel AND #sSst AND NOT #iStartFrmFibroseq;
END_REGION

REGION Network 74: STATE Num:100 Wait For Start Low
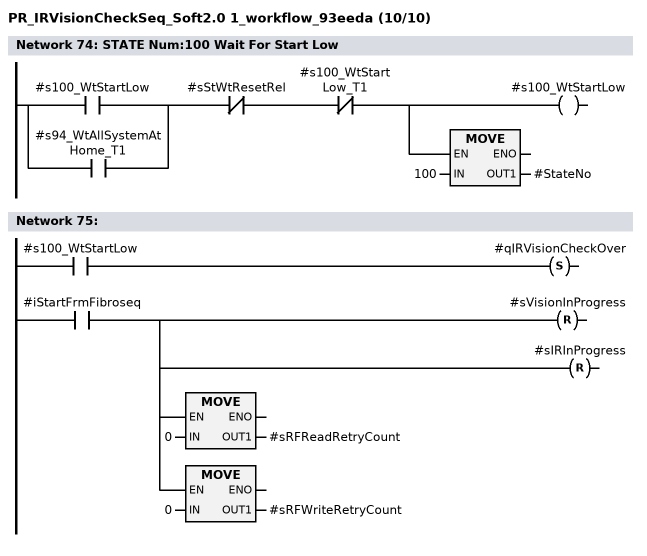
   RUNG wire#powerrail
      Contact( #s100_WtStartLow )
      wire#w1
      I_Contact( #sStWtResetRel )
      I_Contact( #s100_WtStartLow_T1 )
      wire#w2
      Coil( #s100_WtStartLow )
   END_RUNG
   RUNG wire#powerrail
      Contact( #s94_WtAllSystemAtHome_T1 )
   END_RUNG wire#w1
   RUNG wire#w2
      { S7_GenerateENO := "TRUE" } Move(in := 100, out1 => #StateNo)
   END_RUNG
   // the same network as SCL:
   #s100_WtStartLow := (#s100_WtStartLow OR #s94_WtAllSystemAtHome_T1) AND NOT #sStWtResetRel AND NOT #s100_WtStartLow_T1;
   IF #s100_WtStartLow THEN #StateNo := 100; END_IF;
END_REGION

REGION Network 75
   RUNG wire#powerrail
      Contact( #s100_WtStartLow )
      S_Coil( #qIRVisionCheckOver )
   END_RUNG
   RUNG wire#powerrail
      Contact( #iStartFrmFibroseq )
      wire#w1
      R_Coil( #sVisionInProgress )
   END_RUNG
   RUNG wire#w1
      R_Coil( #sIRInProgress )
   END_RUNG
   RUNG wire#w1
      Move(in := 0, out1 => #sRFReadRetryCount)
   END_RUNG
   RUNG wire#w1
      Move(in := 0, out1 => #sRFWriteRetryCount)
   END_RUNG
   // the same network as SCL:
   IF #s100_WtStartLow THEN #qIRVisionCheckOver := TRUE; END_IF;
   IF #iStartFrmFibroseq THEN
       #sVisionInProgress := FALSE;
       #sIRInProgress := FALSE;
       #sRFReadRetryCount := 0;
       #sRFWriteRetryCount := 0;
   END_IF;
END_REGION
END_FUNCTION_BLOCK
